(* IEC 61131-3 sources: rusty/compiler/plc_cfc/fixtures/blocks/valid/generic_chain, 1 file *)

(* ---- myGenAdd.st ---- *)
FUNCTION myGenAdd<T: ANY_NUM> : T
VAR_INPUT
    a : T;
    b : T;
END_VAR
END_FUNCTION

FUNCTION myGenAdd__INT : INT
VAR_INPUT
    a : INT;
    b : INT;
END_VAR
    myGenAdd__INT := a + b;
END_FUNCTION

FUNCTION myGenAdd__DINT : DINT
VAR_INPUT
    a : DINT;
    b : DINT;
END_VAR
    myGenAdd__DINT := a + b;
END_FUNCTION
